(* IEC 61131-3 sources: llm-plc-st-eval/data/processed_v2/gpt-4o/I5/zero_shot, 3 files *)

(* ---- ejec_1.st ---- *)
FUNCTION_BLOCK FB_Clasificadora
VAR_INPUT
    sensorPresencia : BOOL;  // Sensor que detecta la presencia de una pieza
    sensorAltura : BOOL;     // Sensor que detecta si la pieza es alta
END_VAR

VAR_OUTPUT
    banda : BOOL;            // Salida para activar la banda transportadora
    piston : BOOL;           // Salida para activar el pistón desviador
    nAltas : INT;            // Contador de piezas altas
    nBajas : INT;            // Contador de piezas bajas
END_VAR

VAR
    estado : INT;            // Estado del sistema
    temporizadorDesvio : TON; // Temporizador para el retraso del pistón
    temporizadorPiston : TON; // Temporizador para la duración del pistón
END_VAR

// Inicialización
banda := TRUE; // La banda siempre está activa

// Máquina de estados para el control del pistón y conteo
CASE estado OF
    0: // Estado de espera
        IF sensorPresencia THEN
            IF sensorAltura THEN
                // La pieza es alta, iniciar temporizador de desvío
                temporizadorDesvio(IN := TRUE, PT := T#2S);
                estado := 1;
            ELSE
                // La pieza es baja, incrementar contador de bajas
                nBajas := nBajas + 1;
            END_IF;
        END_IF;

    1: // Esperando el tiempo de desvío
        IF temporizadorDesvio.Q THEN
            // Activar pistón y temporizador de pistón
            piston := TRUE;
            temporizadorPiston(IN := TRUE, PT := T#1S);
            estado := 2;
        END_IF;

    2: // Pistón activado
        IF temporizadorPiston.Q THEN
            // Desactivar pistón y resetear temporizadores
            piston := FALSE;
            temporizadorDesvio(IN := FALSE);
            temporizadorPiston(IN := FALSE);
            // Incrementar contador de altas
            nAltas := nAltas + 1;
            estado := 0;
        END_IF;
END_CASE;
END_FUNCTION_BLOCK

(* ---- ejec_2.st ---- *)
FUNCTION_BLOCK FB_Clasificadora
VAR_INPUT
    sensorPresencia : BOOL;  // Sensor que detecta la presencia de una pieza
    sensorAltura : BOOL;     // Sensor que detecta si la pieza es alta
END_VAR

VAR_OUTPUT
    banda : BOOL;            // Salida para activar la banda transportadora
    piston : BOOL;           // Salida para activar el pistón desviador
    nAltas : INT;            // Contador de piezas altas
    nBajas : INT;            // Contador de piezas bajas
END_VAR

VAR
    estado : INT;            // Estado del sistema
    temporizadorDesvio : TON; // Temporizador para el retraso de 2 segundos
    temporizadorPiston : TON; // Temporizador para la duración de 1 segundo del pistón
    piezaAltaDetectada : BOOL; // Indica si se detectó una pieza alta
END_VAR

// Inicialización
banda := TRUE; // La banda siempre está activa

// Máquina de estados para el control del pistón y conteo de piezas
CASE estado OF
    0: // Estado inicial, esperando detección de pieza
        IF sensorPresencia THEN
            IF sensorAltura THEN
                piezaAltaDetectada := TRUE;
                temporizadorDesvio(IN := TRUE, PT := T#2S);
            ELSE
                nBajas := nBajas + 1;
            END_IF;
            estado := 1;
        END_IF;

    1: // Esperando el tiempo de retraso para activar el pistón
        temporizadorDesvio(IN := sensorPresencia AND piezaAltaDetectada);
        IF temporizadorDesvio.Q THEN
            piston := TRUE;
            temporizadorPiston(IN := TRUE, PT := T#1S);
            estado := 2;
        END_IF;

    2: // Activando el pistón durante 1 segundo
        temporizadorPiston(IN := TRUE);
        IF temporizadorPiston.Q THEN
            piston := FALSE;
            nAltas := nAltas + 1;
            piezaAltaDetectada := FALSE;
            estado := 0;
        END_IF;
END_CASE;
END_FUNCTION_BLOCK

(* ---- ejec_3.st ---- *)
FUNCTION_BLOCK FB_Clasificadora
VAR_INPUT
    sensorPresencia : BOOL; // Sensor que detecta la presencia de una pieza
    sensorAltura : BOOL;    // Sensor que detecta si la pieza es alta
END_VAR

VAR_OUTPUT
    banda : BOOL;   // Control de la banda transportadora
    piston : BOOL;  // Control del pistón desviador
    nAltas : INT;   // Contador de piezas altas
    nBajas : INT;   // Contador de piezas bajas
END_VAR

VAR
    estado : INT;           // Estado del proceso
    temporizador : TON;     // Temporizador para el retraso del pistón
    activarPiston : BOOL;   // Señal para activar el pistón
END_VAR

// Inicialización
banda := TRUE; // La banda siempre está activa

// Máquina de estados para el control del proceso
CASE estado OF
    0: // Estado inicial
        IF sensorPresencia THEN
            IF sensorAltura THEN
                // La pieza es alta, iniciar temporizador para el pistón
                temporizador(IN := TRUE, PT := T#2S);
                estado := 1;
            ELSE
                // La pieza es baja, incrementar contador
                nBajas := nBajas + 1;
                estado := 0; // Volver al estado inicial
            END_IF
        END_IF

    1: // Esperar 2 segundos para activar el pistón
        temporizador(IN := TRUE, PT := T#2S);
        IF temporizador.Q THEN
            // Activar el pistón por 1 segundo
            activarPiston := TRUE;
            temporizador(IN := FALSE);
            temporizador(IN := TRUE, PT := T#1S);
            estado := 2;
        END_IF

    2: // Mantener el pistón activado por 1 segundo
        piston := activarPiston;
        IF temporizador.Q THEN
            // Desactivar el pistón y actualizar contador
            activarPiston := FALSE;
            piston := FALSE;
            nAltas := nAltas + 1;
            estado := 0; // Volver al estado inicial
        END_IF
END_CASE
END_FUNCTION_BLOCK
